Fanuc KAREL source: kt00747.KL

-- PROVISIONAL review KL for V1013-1; original PC SHA256 b8550907dbec4d93489ffb4da1c1a50f9c77f1b86daa2420dc9647ee2cb3b3a2
-- Incomplete behavior may be omitted. Consult companion uncertainty JSON. Do not deploy.
PROGRAM KT00747
%NOLOCKGROUP
BEGIN
  -- UNRESOLVED_PC offsets 5-18; opcodes 22,1D,23
  -- UNRESOLVED_PC offsets 23-27; opcodes 7F
END KT00747
